(*
SPDX-FileCopyrightText: © 2026 Oleksandr Tiutyk <trofimich@gmail.com>
SPDX-License-Identifier: MIT
License: https://opensource.org/license/mit
*)

(*!
<summary>Groups timer timing, lifecycle and restart scenarios.</summary>
<description>
Owns the test cases and their fixed child array. Use from a single PLC task and keep the group at a stable address.
</description>
*)

{attribute 'no_assign'}
{attribute 'no_explicit_call' := 'do not call this function block directly'}
FUNCTION_BLOCK TimerTimingTestGroup EXTENDS TOF_Testing.TestGroup<13>
VAR_STAT
	{attribute 'hide'}
	_ClassName : STRING := __POUNAME();
END_VAR
VAR
	_PositiveIntervalSameCallRestart : TimerCompletionPulseTest(
		name := "PositiveIntervalSameCallRestart",
		parent := THIS^,
		interval := T#30MS
	);
	_ZeroIntervalSameCallRestart : TimerCompletionPulseTest(
		name := "ZeroIntervalSameCallRestart",
		parent := THIS^,
		interval := TOF_Core.Times.MIN_VALUE
	);
	_DefaultNameAndMetadata : TimerMetadataTest(
		name := "DefaultNameAndMetadata",
		parent := THIS^
	);
	_CancelBeforeFirstExecuteAndReuse : TimerCancelBeforeExecuteTest(
		name := "CancelBeforeFirstExecuteAndReuse",
		parent := THIS^
	);
	_ResetAfterCompletion : TimerResetAfterCompletionTest(
		name := "ResetAfterCompletion",
		parent := THIS^
	);
	_IntervalAssignmentPreservesObservation : TimerIntervalObservationTest(
		name := "IntervalAssignmentPreservesObservation",
		parent := THIS^
	);
	_RestartWaitsForStopping : TimerPendingRestartTest(
		name := "RestartWaitsForStopping",
		parent := THIS^
	);
	_RestartPreservesIntervalOnResetFailure : TimerRestartResetFailureTest(
		name := "RestartPreservesIntervalOnResetFailure",
		parent := THIS^
	);
	_RestartRetainsIntervalOnStartFailure : TimerRestartStartFailureTest(
		name := "RestartRetainsIntervalOnStartFailure",
		parent := THIS^
	);
	_CompletionCallbackCanReset : TimerCompletionCallbackTest(
		name := "CompletionCallbackCanReset",
		parent := THIS^
	);
	_DelayedFirstExecuteUsesStartAnchor : DelayedTimerObservationTest(
		name := "DelayedFirstExecuteUsesStartAnchor",
		parent := THIS^,
		scenario := DELAYED_TIMER_TEST_SCENARIO.AFTER_START
	);
	_CancelAfterUnobservedExpiry : DelayedTimerObservationTest(
		name := "CancelAfterUnobservedExpiry",
		parent := THIS^,
		scenario := DELAYED_TIMER_TEST_SCENARIO.CANCEL_BEFORE_EXECUTE
	);
	_PositiveRestartUsesStartAnchor : DelayedTimerObservationTest(
		name := "PositiveRestartUsesStartAnchor",
		parent := THIS^,
		scenario := DELAYED_TIMER_TEST_SCENARIO.AFTER_ACTIVE_RESTART
	);

	_Children : ARRAY [0.._ChildCount - 1] OF TOF_Testing.ITestElement :=
	[
		_PositiveIntervalSameCallRestart,
		_ZeroIntervalSameCallRestart,
		_DefaultNameAndMetadata,
		_CancelBeforeFirstExecuteAndReuse,
		_ResetAfterCompletion,
		_IntervalAssignmentPreservesObservation,
		_RestartWaitsForStopping,
		_RestartPreservesIntervalOnResetFailure,
		_RestartRetainsIntervalOnStartFailure,
		_CompletionCallbackCanReset,
		_DelayedFirstExecuteUsesStartAnchor,
		_CancelAfterUnobservedExpiry,
		_PositiveRestartUsesStartAnchor
	];
END_VAR

//! <summary>Borrows the fixed child array. Callers must not modify it.</summary>
{attribute 'monitoring' := 'call'}
PROPERTY Children : REFERENCE TO ARRAY [0.._ChildCount - 1] OF TOF_Testing.ITestElement
GET
Children REF= _Children;
END_GET
END_PROPERTY

//! <summary>Borrows the concrete class name. Callers must not modify it.</summary>
{attribute 'monitoring' := 'call'}
PROPERTY ClassName : REFERENCE TO STRING
GET
ClassName REF= _ClassName;
END_GET
END_PROPERTY

//! <summary>Borrows the compiler-initialized namespace. Callers must not modify it.</summary>
{attribute 'monitoring' := 'call'}
PROPERTY NamespaceName : REFERENCE TO STRING
GET
NamespaceName REF= CurrentNamespace.Name;
END_GET
END_PROPERTY

//! <summary>Reports the concrete instance size in bytes.</summary>
{attribute 'monitoring' := 'call'}
PROPERTY SelfSize : ULINT
GET
SelfSize := XSIZEOF(THIS^);
END_GET
END_PROPERTY

END_FUNCTION_BLOCK

(* stored: Version 1.1.0.1
   POU TimerTimingTestGroup: Id {2d83cb3b-db5c-454f-b332-d9149d0e7435}, SpecialFunc None
   Property Children: Id {6f4de77e-ca97-4535-8cfe-6e77de1377be}
   Get Get: Id {fe4bb99c-9245-4019-b253-80ec5ef187ae}
   Property ClassName: Id {ea83f2fe-8ee4-42ef-b386-9bbe7ba5f0b2}
   Get Get: Id {5e7c2296-c41d-49ed-9f9d-301d1fc0e57e}
   Property NamespaceName: Id {1245437d-7444-4c03-af0c-8c68d493dc0d}
   Get Get: Id {461005d0-ec78-4783-ac77-83b7de983acd}
   Property SelfSize: Id {7e712336-255f-40fc-803c-44d0976e682f}
   Get Get: Id {0d50a699-6150-4633-b203-d62d0c40109b} *)
